// TIA Portal V18 export
DATA_BLOCK "DB_MB_RTU_MasterConfig"   // DB10
{ S7_Optimized_Access := 'TRUE' }
// stored: MemoryReserve 0
   VAR
      REQ : Bool;
      MB_ADDR : UInt := 1;
      MODE : USInt;
      DATA_ADDR : UDInt;
      DATA_LEN : UInt;
      DONE : Bool;
      BUSY : Bool;
      ERROR : Bool;
      STATUS : Word;
      ptrAddr : Int;
      "Step" : Int;
      StepRequest : Int;
   END_VAR
BEGIN
END_DATA_BLOCK
